// TIA Portal V19 export
DATA_BLOCK "G120XA_DATA"   // DB92
{ S7_Optimized_Access := 'FALSE' }
   VAR RETAIN
      COLD_SKID_CP01 : Struct
         START_CMD : Bool;
         FAULT_RESET : Bool;
         RUN_FBK : Bool;
         TRIP_FBK : Bool;
         SPEED_REF : Int;
         ACT_SPEED : Int;
      END_STRUCT;
      COLD_SKID_CP02 : Struct
         START_CMD : Bool;
         FAULT_RESET : Bool;
         RUN_FBK : Bool;
         TRIP_FBK : Bool;
         SPEED_REF : Int;
         ACT_SPEED : Int;
      END_STRUCT;
      COLD_SKID_CP03 : Struct
         START_CMD : Bool;
         FAULT_RESET : Bool;
         RUN_FBK : Bool;
         TRIP_FBK : Bool;
         SPEED_REF : Int;
         ACT_SPEED : Int;
      END_STRUCT;
      COLD_SKID_DRIVE_CMD : Int;
      COLD_SKID_DRIVE_FBK : Int;
      "A/m" : Int;
   END_VAR
BEGIN
END_DATA_BLOCK
